// TIA Portal V19 export
ORGANIZATION_BLOCK "Cyclic1s"   // OB31, FBD, CyclicInterrupt
{ S7_Optimized_Access := 'TRUE' }
// stored: SetENOAutomatically false
   VAR_INPUT
      Initial_Call : Bool;   // Initial call of this OB
      Event_Count : Int;   // Events discarded
   END_VAR
BEGIN

REGION Network 1
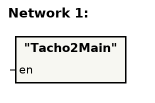
   "Tacho2Main"();
END_REGION
END_ORGANIZATION_BLOCK
